Fanuc KAREL source: KX00017.KL

PROGRAM KX00017
%NOLOCKGROUP
VAR
  I: INTEGER
  J: INTEGER
  B: BOOLEAN
  F: FILE
  S: STRING[80]
  P: XYZWPR
BEGIN
  WAIT FOR DIN[2]
END KX00017
